Omron Sysmac Studio project 자동화산업기사-고건우_3 (Sysmac Studio 1.53.0.9, StandardProject)

# Controller CPU1: NX102-1020 version 1.33
Units and slaves: 노드1 : NX-ECC203 (E001); 유니트 1 : NX-ID6142-6 (N1); 유니트 2 : NX-OD6121-6 (N2); 유니트 1 : NX-PF0730 (N3); 유니트 2 : NX-ILM400 (N4); 유니트 4 : NX-SID800 (N6); 유니트 5 : NX-SOD400 (N7)
Task PrimaryTask (priority 4, period or condition 2000): Program0

TYPE D_out : UNION
    dw : DWORD;
    b : ARRAY[0..32] OF bool;
END_UNION END_TYPE
TYPE D_in : UNION
    dw : DWORD;
    b : ARRAY[0..32] OF bool;
END_UNION END_TYPE
TYPE U_IO16 : UNION
    W : WORD;
    B : ARRAY[1..32] OF BOOL;
END_UNION END_TYPE
TYPE S_RobotIO : STRUCT
    IO : U_IO16;
END_STRUCT END_TYPE

VAR_GLOBAL
    Bot_Task_Pause : BOOL;  (* 로봇 - 테스크 일시정지; at ECAT://node#[1,2]/Output Bit 32 bits/Output Bit 04 *)
    Discharge_F_SOL : BOOL;  (* at ECAT://node#[1,2]/Output Bit 32 bits/Output Bit 05 *)
    Discharge_R_SS : BOOL;  (* at ECAT://node#[1,1]/Input Bit 32 bits/Input Bit 25 *)
    N1_Input_Bit_26 : BOOL;
    N1_Input_Bit_27 : BOOL;
    N1_Input_Bit_28 : BOOL;
    N1_Input_Bit_29 : BOOL;
    N1_Input_Bit_30 : BOOL;
    N1_Input_Bit_31 : BOOL;
    MotM : WORD;  (* at ECAT://node#2/Command *)
    Vision_Trigger : BOOL;  (* at ECAT://node#4/Line0 Trigger *)
    MotM_Status : WORD;  (* at ECAT://node#2/Status *)
    Robot_Recv : S_RobotIO;
    Robot_Send : S_RobotIO;
    Robot_In : ARRAY[0..237] OF WORD;  (* network input *)
    Robot_Out : ARRAY[0..105] OF WORD;  (* network output *)
END_VAR
VAR_GLOBAL RETAIN
    Bot_IO : ARRAY[1..7] OF WORD := [16#01, 16#02, 16#04, 16#08, 16#10, 16#20, 16#40];
END_VAR
VAR_GLOBAL
    Discharge_R_SOL : BOOL;  (* at ECAT://node#[1,2]/Output Bit 32 bits/Output Bit 06 *)
    Bot_Task_Stop : BOOL;  (* 로봇 - 프로그램 정지; at ECAT://node#[1,2]/Output Bit 32 bits/Output Bit 24 *)
    TWL_R : BOOL;  (* 타워램프 - RED; at ECAT://node#[1,2]/Output Bit 32 bits/Output Bit 20 *)
    TWL_Y : BOOL;  (* 타워램프 - YELLOW; at ECAT://node#[1,2]/Output Bit 32 bits/Output Bit 21 *)
    TWL_G : BOOL;  (* 타워램프 - GREEN; at ECAT://node#[1,2]/Output Bit 32 bits/Output Bit 22 *)
    Bot_Task_ON : BOOL;  (* 로봇 - 태스크 실행; at ECAT://node#[1,2]/Output Bit 32 bits/Output Bit 23 *)
    Vision_SS : BOOL;  (* at ECAT://node#[1,1]/Input Bit 32 bits/Input Bit 19 *)
    Stopper_SS : BOOL;  (* at ECAT://node#[1,1]/Input Bit 32 bits/Input Bit 24 *)
    Magazine_SS : BOOL;  (* at ECAT://node#[1,1]/Input Bit 32 bits/Input Bit 23 *)
    Discharge_F_SS : BOOL;  (* at ECAT://node#[1,1]/Input Bit 32 bits/Input Bit 26 *)
    Bot_Task_Resume : BOOL;  (* 로봇 - 테스크 재개; at ECAT://node#[1,2]/Output Bit 32 bits/Output Bit 13 *)
    Vis_Data : DINT;  (* at ECAT://node#4/Line0 DINT Result Data 0 *)
    H_Count_Val : INT;
    H_Total_Val : INT;
    Robot_DI : S_RobotIO;
    MultiMode_PB : BOOL;
    SingleMode_PB : BOOL;
    Target_Slot_Status : ARRAY[1..6] OF BOOL;
    Stop_PB : BOOL;
    Auto_PB : BOOL;
    Manual_PB : BOOL;
    MotMV_PB : BOOL;
    MotST_PB : BOOL;
    F_SOL_PB : BOOL;
    R_SOL_PB : BOOL;
    Clamp_PB : BOOL;
    UnClamp_PB : BOOL;
    H_Err_Val : INT;
    Auto_Busy : BOOL;
    Manual_Busy : BOOL;
    Pause_PB : BOOL;
    Resume_PB : BOOL;
    Estop_PB : BOOL;
    RST_PB : BOOL;
    gDMemory : WORD;
END_VAR

(* Program Program0: safety or other program stored in binary form, left out *)

PROGRAM Program0
VAR
    i : INT;
    Start : BOOL;
    Vis_ON : BOOL;
    data : INT;
    Sensor_OK : BOOL;
    Pause : BOOL;
    T0 : TON;
    T0TImer : DINT;
    TP0 : TP;
    AT0 : AccumulationTimer;
    Auto : Equipment;
END_VAR
VAR_EXTERNAL
    MotM : WORD;
    Vision_Trigger : BOOL;
    MotM_Status : WORD;
    Magazine_SS : BOOL;
    Discharge_R_SS : BOOL;
    Stopper_SS : BOOL;
    Discharge_F_SS : BOOL;
    Vision_SS : BOOL;
    Vis_Data : DINT;
    Robot_Recv : S_RobotIO;
    Discharge_F_SOL : BOOL;
    Discharge_R_SOL : BOOL;
    Robot_Send : S_RobotIO;
    Bot_Task_Stop : BOOL;
    Bot_Task_ON : BOOL;
    Robot_In : ARRAY[0..237] OF WORD;
    Robot_Out : ARRAY[0..105] OF WORD;
    Bot_Task_Pause : BOOL;
    Bot_Task_Resume : BOOL;
    Bot_IO : ARRAY[1..7] OF WORD;
    H_Count_Val : INT;
    H_Total_Val : INT;
    Robot_DI : S_RobotIO;
    MultiMode_PB : BOOL;
    SingleMode_PB : BOOL;
    Target_Slot_Status : ARRAY[1..6] OF BOOL;
    Stop_PB : BOOL;
    Auto_PB : BOOL;
    Manual_PB : BOOL;
    MotMV_PB : BOOL;
    MotST_PB : BOOL;
    F_SOL_PB : BOOL;
    R_SOL_PB : BOOL;
    Clamp_PB : BOOL;
    UnClamp_PB : BOOL;
    H_Err_Val : INT;
    Auto_Busy : BOOL;
    Manual_Busy : BOOL;
    Pause_PB : BOOL;
    Resume_PB : BOOL;
    Estop_PB : BOOL;
    RST_PB : BOOL;
    TWL_G : BOOL;
    TWL_R : BOOL;
    TWL_Y : BOOL;
END_VAR

(* Section Section0: ladder, written here as Structured Text *)

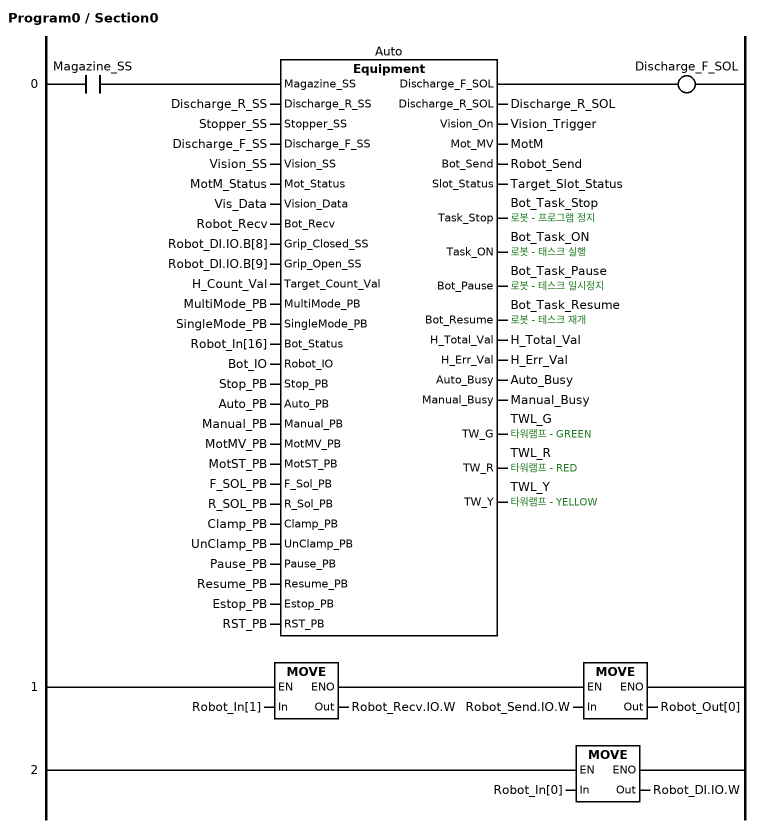
(* Rung 0 *)
Auto(Magazine_SS := Magazine_SS, Discharge_R_SS := Discharge_R_SS, Stopper_SS := Stopper_SS, Discharge_F_SS := Discharge_F_SS, Vision_SS := Vision_SS, Mot_Status := MotM_Status, Vision_Data := Vis_Data, Bot_Recv := Robot_Recv, Grip_Closed_SS := Robot_DI.IO.B[8], Grip_Open_SS := Robot_DI.IO.B[9], Target_Count_Val := H_Count_Val, MultiMode_PB := MultiMode_PB, SingleMode_PB := SingleMode_PB, Bot_Status := Robot_In[16], Robot_IO := Bot_IO, Stop_PB := Stop_PB, Auto_PB := Auto_PB, Manual_PB := Manual_PB, MotMV_PB := MotMV_PB, MotST_PB := MotST_PB, F_Sol_PB := F_SOL_PB, R_Sol_PB := R_SOL_PB, Clamp_PB := Clamp_PB, UnClamp_PB := UnClamp_PB, Pause_PB := Pause_PB, Resume_PB := Resume_PB, Estop_PB := Estop_PB, RST_PB := RST_PB, Discharge_R_SOL => Discharge_R_SOL, Vision_On => Vision_Trigger, Mot_MV => MotM, Bot_Send => Robot_Send, Slot_Status => Target_Slot_Status, Task_Stop => Bot_Task_Stop, Task_ON => Bot_Task_ON, Bot_Pause => Bot_Task_Pause, Bot_Resume => Bot_Task_Resume, H_Total_Val => H_Total_Val, H_Err_Val => H_Err_Val, Auto_Busy => Auto_Busy, Manual_Busy => Manual_Busy, TW_G => TWL_G, TW_R => TWL_R, TW_Y => TWL_Y);
Discharge_F_SOL := Auto.Discharge_F_SOL;
(* Rung 1 *)
Robot_Recv.IO.W := Robot_In[1];
Robot_Out[0] := Robot_Send.IO.W;
(* Rung 2 *)
Robot_DI.IO.W := Robot_In[0];
END_PROGRAM

FUNCTION_BLOCK MPS
VAR
    data : INT;
    T0 : TON;
END_VAR
VAR_INPUT
    MPS_Start : BOOL;
    Discharge_R_SS : BOOL;
    Stopper_SS : BOOL;
END_VAR
VAR_OUTPUT
    Discharge_F_SOL : BOOL;
END_VAR
VAR_INPUT
    Discharge_F_SS : BOOL;
END_VAR
VAR_OUTPUT
    Discharge_R_SOL : BOOL;
END_VAR
VAR_INPUT
    Vision_SS : BOOL;
END_VAR
VAR_OUTPUT
    Vision_On : BOOL;
END_VAR
VAR_INPUT
    Mot_Status : WORD;
END_VAR
VAR_OUTPUT
    MPS_Done : BOOL;
END_VAR
VAR_INPUT
    Cmd_Ack : BOOL;
END_VAR
VAR_OUTPUT
    MPS_Busy : BOOL;
END_VAR
VAR_INPUT
    Vision_Data : DINT;
END_VAR
VAR_OUTPUT
    VIs_NO : DINT;
END_VAR
VAR_IN_OUT
    Mot_MV : WORD;
END_VAR
VAR_INPUT
    Estop_Active : BOOL;
    RST_Active : BOOL;
    Slot_Status : ARRAY[1..6] OF BOOL;
    Pause_Active : BOOL;
END_VAR
VAR
    _e1 : R_TRIG;
    _p2 : BOOL;
    _p3 : BOOL;
END_VAR
(* ladder, written here as Structured Text *)

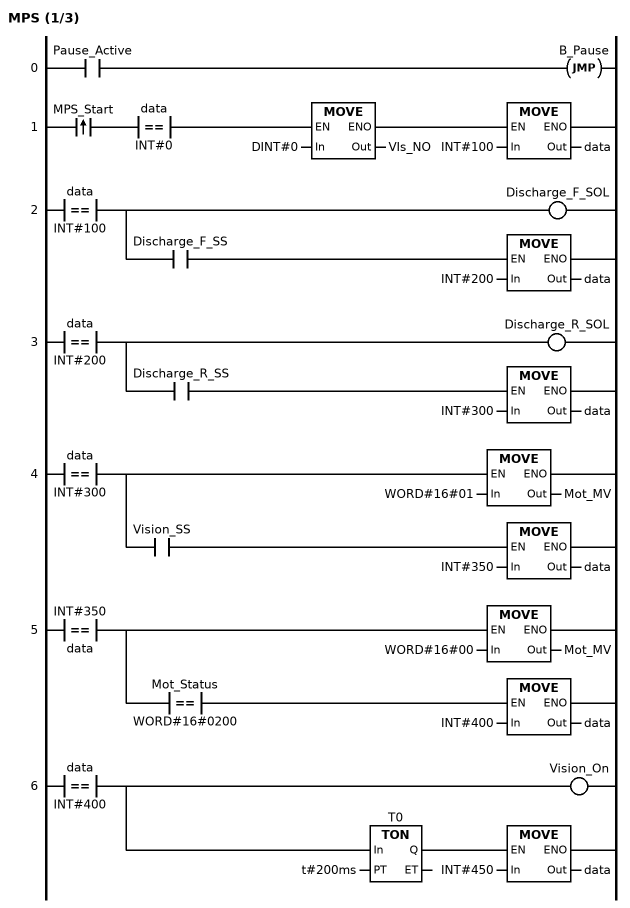
(* Rung 0 *)
IF Pause_Active THEN JMP B_Pause; END_IF;
(* Rung 1 *)
_e1(CLK := MPS_Start);
IF _e1.Q AND (data = INT#0) THEN
    VIs_NO := DINT#0;
    data := INT#100;
END_IF;
(* Rung 2 *)
Discharge_F_SOL := data = INT#100;
IF (data = INT#100) AND Discharge_F_SS THEN data := INT#200; END_IF;
(* Rung 3 *)
Discharge_R_SOL := data = INT#200;
IF (data = INT#200) AND Discharge_R_SS THEN data := INT#300; END_IF;
(* Rung 4 *)
IF data = INT#300 THEN Mot_MV := WORD#16#01; END_IF;
IF (data = INT#300) AND Vision_SS THEN data := INT#350; END_IF;
(* Rung 5 *)
IF INT#350 = data THEN Mot_MV := WORD#16#00; END_IF;
IF (INT#350 = data) AND (Mot_Status = WORD#16#0200) THEN data := INT#400; END_IF;
(* Rung 6 *)
Vision_On := data = INT#400;
T0(In := data = INT#400, PT := t#200ms);
IF T0.Q THEN data := INT#450; END_IF;

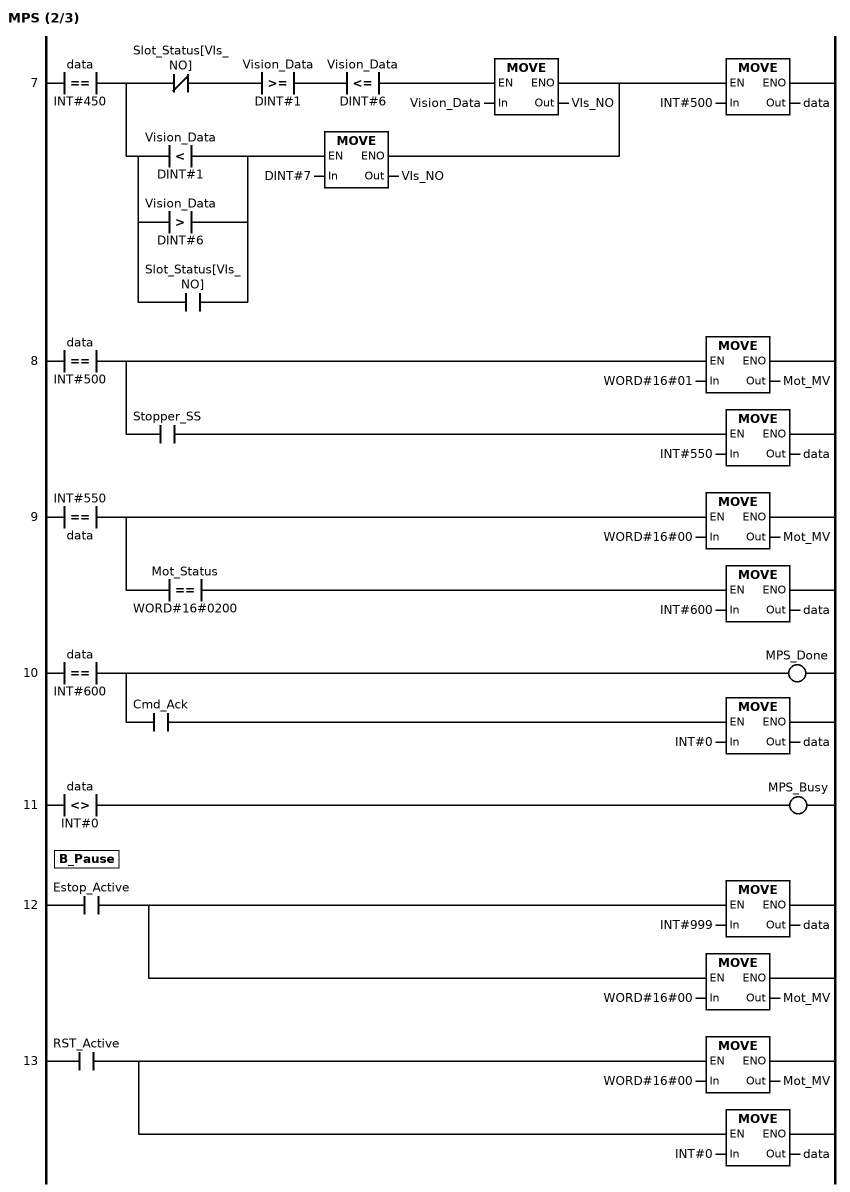
(* Rung 7 *)
_p2 := (data = INT#450) AND NOT Slot_Status[VIs_NO] AND (Vision_Data >= DINT#1) AND (Vision_Data <= DINT#6);
IF _p2 THEN VIs_NO := Vision_Data; END_IF;
_p3 := (data = INT#450) AND ((Vision_Data < DINT#1) OR (Vision_Data > DINT#6) OR Slot_Status[VIs_NO]);
IF _p3 THEN VIs_NO := DINT#7; END_IF;
IF _p2 OR _p3 THEN data := INT#500; END_IF;
(* Rung 8 *)
IF data = INT#500 THEN Mot_MV := WORD#16#01; END_IF;
IF (data = INT#500) AND Stopper_SS THEN data := INT#550; END_IF;
(* Rung 9 *)
IF INT#550 = data THEN Mot_MV := WORD#16#00; END_IF;
IF (INT#550 = data) AND (Mot_Status = WORD#16#0200) THEN data := INT#600; END_IF;
(* Rung 10 *)
MPS_Done := data = INT#600;
IF (data = INT#600) AND Cmd_Ack THEN data := INT#0; END_IF;
(* Rung 11 *)
MPS_Busy := data <> INT#0;
(* Rung 12 *)
B_Pause:
IF Estop_Active THEN
    data := INT#999;
    Mot_MV := WORD#16#00;
END_IF;
(* Rung 13 *)
IF RST_Active THEN
    Mot_MV := WORD#16#00;
    data := INT#0;
END_IF;

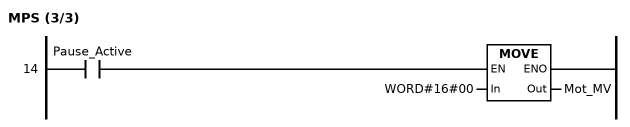
(* Rung 14 *)
IF Pause_Active THEN Mot_MV := WORD#16#00; END_IF;
END_FUNCTION_BLOCK

FUNCTION_BLOCK Robot
VAR
    data : INT;
    T0 : TON;
END_VAR
VAR_INPUT
    Bot_Start : BOOL;
END_VAR
VAR_OUTPUT
    Bot_Done : BOOL;
    Bot_Busy : BOOL;
END_VAR
VAR_IN_OUT
    Slot_Status : ARRAY[1..6] OF BOOL;
END_VAR
VAR_INPUT
    Estop_Active : BOOL;
    RST_Active : BOOL;
    Pause_Active : BOOL;
    Target_Slot_No : DINT;
    MultiMode : BOOL;
END_VAR
VAR_IN_OUT
    Bot_Send : S_RobotIO;
END_VAR
VAR_INPUT
    Bot_Recv : S_RobotIO;
    Bot_Status : WORD;
    Bot_IO : ARRAY[1..7] OF WORD;
END_VAR
VAR_IN_OUT
    H_Total_Val : INT;
    H_Err_Val : INT;
END_VAR
VAR
    _p1 : BOOL;
    _e2 : R_TRIG;
    _e3 : R_TRIG;
END_VAR
(* ladder, written here as Structured Text *)

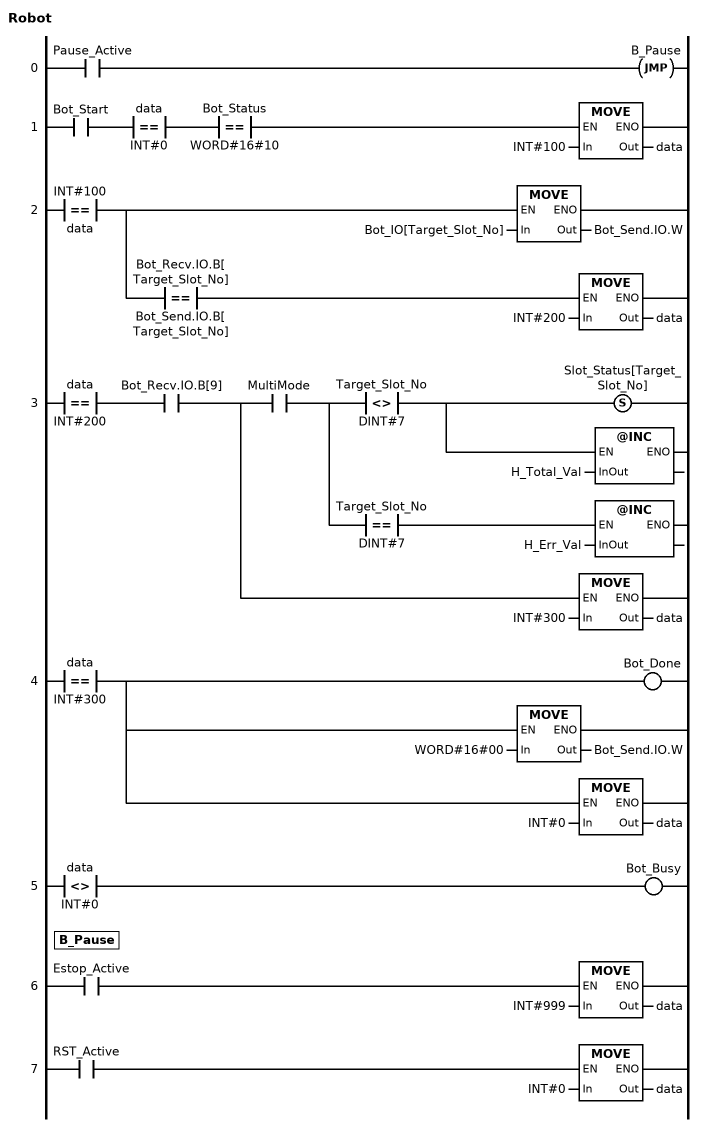
(* Rung 0 *)
IF Pause_Active THEN JMP B_Pause; END_IF;
(* Rung 1 *)
IF Bot_Start AND (data = INT#0) AND (Bot_Status = WORD#16#10) THEN data := INT#100; END_IF;
(* Rung 2 *)
IF INT#100 = data THEN Bot_Send.IO.W := Bot_IO[Target_Slot_No]; END_IF;
IF (INT#100 = data) AND (Bot_Recv.IO.B[Target_Slot_No] = Bot_Send.IO.B[Target_Slot_No]) THEN
    data := INT#200;
END_IF;
(* Rung 3 *)
_p1 := (data = INT#200) AND Bot_Recv.IO.B[9] AND MultiMode;
IF _p1 AND (Target_Slot_No <> DINT#7) THEN Slot_Status[Target_Slot_No] := TRUE; END_IF;
_e2(CLK := _p1 AND (Target_Slot_No <> DINT#7));
IF _e2.Q THEN INC(InOut := H_Total_Val); END_IF;
_e3(CLK := _p1 AND (Target_Slot_No = DINT#7));
IF _e3.Q THEN INC(InOut := H_Err_Val); END_IF;
IF (data = INT#200) AND Bot_Recv.IO.B[9] THEN data := INT#300; END_IF;
(* Rung 4 *)
Bot_Done := data = INT#300;
IF data = INT#300 THEN
    Bot_Send.IO.W := WORD#16#00;
    data := INT#0;
END_IF;
(* Rung 5 *)
Bot_Busy := data <> INT#0;
(* Rung 6 *)
B_Pause:
IF Estop_Active THEN data := INT#999; END_IF;
(* Rung 7 *)
IF RST_Active THEN data := INT#0; END_IF;
END_FUNCTION_BLOCK

FUNCTION_BLOCK Equipment
VAR
    Conveyor : MPS;
    Doosan : Robot;
    Bot_Busy : BOOL;
    Mps_Done : BOOL;
    Mps_Busy : BOOL;
    Vis_No : DINT;
    Bot_Done : BOOL;
    Single_Busy : BOOL;
    Multi_Busy : BOOL;
    C0 : CTU;
    Estop_Active : BOOL;
    RST_Active : BOOL;
    Pause_Active : BOOL;
    Retry : BOOL;
    CTU_RST : BOOL;
    T0 : TON;
    T1 : TON;
    T2 : TON;
    RST_On : BOOL;
    RST_Discharge_R_SOL : BOOL;
    MPS_Discharge_R_SOL : BOOL;
    Stop_Active : BOOL;
    Manual : Passive;
    Manu_Discharge_F_SOL : BOOL;
    Manu_Discharge_R_SOL : BOOL;
    Manu_TWL_G : BOOL;
    MPS_Discharge_F_SOL : BOOL;
    T3 : TON;
    Ready : BOOL;
    Pulse_Pause : BOOL;
    Pause_Eq : BOOL;
END_VAR
VAR_INPUT
    Magazine_SS : BOOL;
    Discharge_R_SS : BOOL;
    Stopper_SS : BOOL;
    Discharge_F_SS : BOOL;
    Vision_SS : BOOL;
    Mot_Status : WORD;
    Vision_Data : DINT;
END_VAR
VAR_OUTPUT
    Discharge_F_SOL : BOOL;
    Discharge_R_SOL : BOOL;
    Vision_On : BOOL;
    Mot_MV : WORD;
END_VAR
VAR_INPUT
    Bot_Recv : S_RobotIO;
END_VAR
VAR_OUTPUT
    Bot_Send : S_RobotIO;
END_VAR
VAR_INPUT
    Grip_Closed_SS : BOOL;
    Grip_Open_SS : BOOL;
END_VAR
VAR_OUTPUT
    Slot_Status : ARRAY[1..6] OF BOOL;
    Task_Stop : BOOL;
END_VAR
VAR_INPUT
    Target_Count_Val : INT;
    MultiMode_PB : BOOL;
    SingleMode_PB : BOOL;
END_VAR
VAR_OUTPUT
    Task_ON : BOOL;
END_VAR
VAR_INPUT
    Bot_Status : WORD;
END_VAR
VAR_OUTPUT
    Bot_Pause : BOOL;
    Bot_Resume : BOOL;
END_VAR
VAR_INPUT
    Robot_IO : ARRAY[1..7] OF WORD;
END_VAR
VAR_OUTPUT
    H_Total_Val : INT;
END_VAR
VAR_INPUT
    Stop_PB : BOOL;
    Auto_PB : BOOL;
    Manual_PB : BOOL;
    MotMV_PB : BOOL;
    MotST_PB : BOOL;
    F_Sol_PB : BOOL;
    R_Sol_PB : BOOL;
    Clamp_PB : BOOL;
    UnClamp_PB : BOOL;
END_VAR
VAR_OUTPUT
    H_Err_Val : INT;
    Auto_Busy : BOOL;
    Manual_Busy : BOOL;
END_VAR
VAR_INPUT
    Pause_PB : BOOL;
    Resume_PB : BOOL;
    Estop_PB : BOOL;
    RST_PB : BOOL;
END_VAR
VAR_OUTPUT
    TW_G : BOOL;
    TW_R : BOOL;
    TW_Y : BOOL;
END_VAR
VAR
    _e1 : R_TRIG;
    _p2 : BOOL;
    _e3 : F_TRIG;
    _e4 : R_TRIG;
    _e5 : R_TRIG;
END_VAR
(* ladder, written here as Structured Text *)

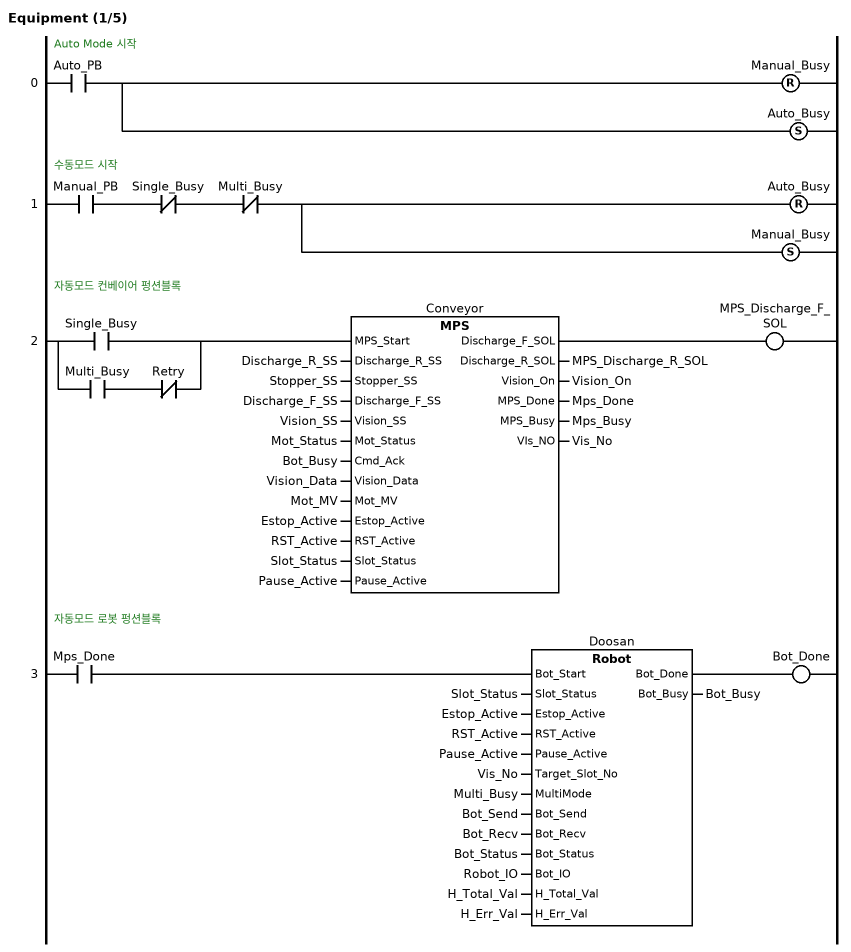
(* Rung 0: Auto Mode 시작 *)
IF Auto_PB THEN
    Manual_Busy := FALSE;
    Auto_Busy := TRUE;
END_IF;
(* Rung 1: 수동모드 시작 *)
IF Manual_PB AND NOT Single_Busy AND NOT Multi_Busy THEN
    Auto_Busy := FALSE;
    Manual_Busy := TRUE;
END_IF;
(* Rung 2: 자동모드 컨베이어 펑션블록 *)
Conveyor(MPS_Start := Single_Busy OR (Multi_Busy AND NOT Retry), Discharge_R_SS := Discharge_R_SS, Stopper_SS := Stopper_SS, Discharge_F_SS := Discharge_F_SS, Vision_SS := Vision_SS, Mot_Status := Mot_Status, Cmd_Ack := Bot_Busy, Vision_Data := Vision_Data, Mot_MV := Mot_MV, Estop_Active := Estop_Active, RST_Active := RST_Active, Slot_Status := Slot_Status, Pause_Active := Pause_Active, Discharge_R_SOL => MPS_Discharge_R_SOL, Vision_On => Vision_On, MPS_Done => Mps_Done, MPS_Busy => Mps_Busy, VIs_NO => Vis_No);
MPS_Discharge_F_SOL := Conveyor.Discharge_F_SOL;
(* Rung 3: 자동모드 로봇 펑션블록 *)
Doosan(Bot_Start := Mps_Done, Slot_Status := Slot_Status, Estop_Active := Estop_Active, RST_Active := RST_Active, Pause_Active := Pause_Active, Target_Slot_No := Vis_No, MultiMode := Multi_Busy, Bot_Send := Bot_Send, Bot_Recv := Bot_Recv, Bot_Status := Bot_Status, Bot_IO := Robot_IO, H_Total_Val := H_Total_Val, H_Err_Val := H_Err_Val, Bot_Busy => Bot_Busy);
Bot_Done := Doosan.Bot_Done;

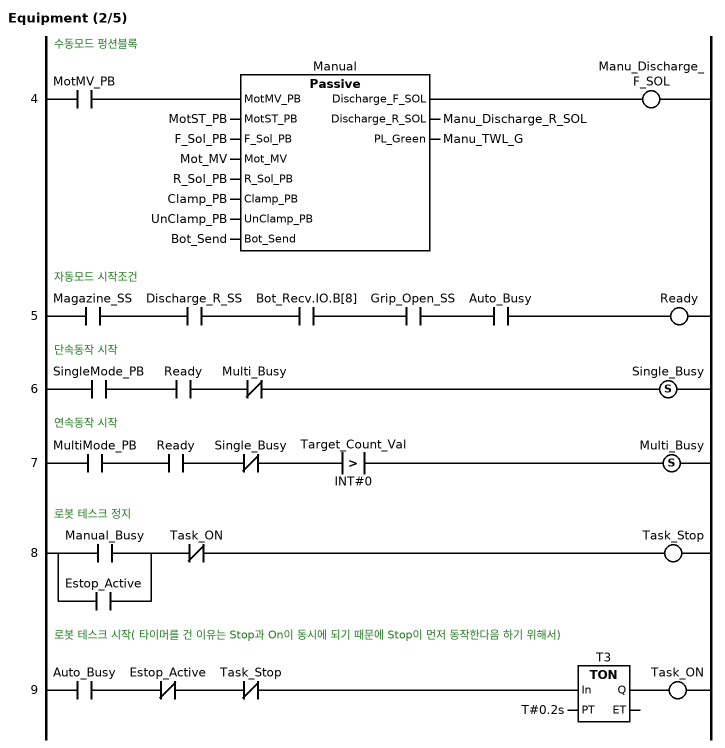
(* Rung 4: 수동모드 펑션블록 *)
Manual(MotMV_PB := MotMV_PB, MotST_PB := MotST_PB, F_Sol_PB := F_Sol_PB, Mot_MV := Mot_MV, R_Sol_PB := R_Sol_PB, Clamp_PB := Clamp_PB, UnClamp_PB := UnClamp_PB, Bot_Send := Bot_Send, Discharge_R_SOL => Manu_Discharge_R_SOL, PL_Green => Manu_TWL_G);
Manu_Discharge_F_SOL := Manual.Discharge_F_SOL;
(* Rung 5: 자동모드 시작조건 *)
Ready := Magazine_SS AND Discharge_R_SS AND Bot_Recv.IO.B[8] AND Grip_Open_SS AND Auto_Busy;
(* Rung 6: 단속동작 시작 *)
IF SingleMode_PB AND Ready AND NOT Multi_Busy THEN Single_Busy := TRUE; END_IF;
(* Rung 7: 연속동작 시작 *)
IF MultiMode_PB AND Ready AND NOT Single_Busy AND (Target_Count_Val > INT#0) THEN
    Multi_Busy := TRUE;
END_IF;
(* Rung 8: 로봇 테스크 정지 *)
Task_Stop := (Manual_Busy OR Estop_Active) AND NOT Task_ON;
(* Rung 9: 로봇 테스크 시작( 타이머를 건 이유는 Stop과 On이 동시에 되기 때문에 Stop이 먼저 동작한다음 하기 위해서) *)
T3(In := Auto_Busy AND NOT Estop_Active AND NOT Task_Stop, PT := T#0.2s);
Task_ON := T3.Q;

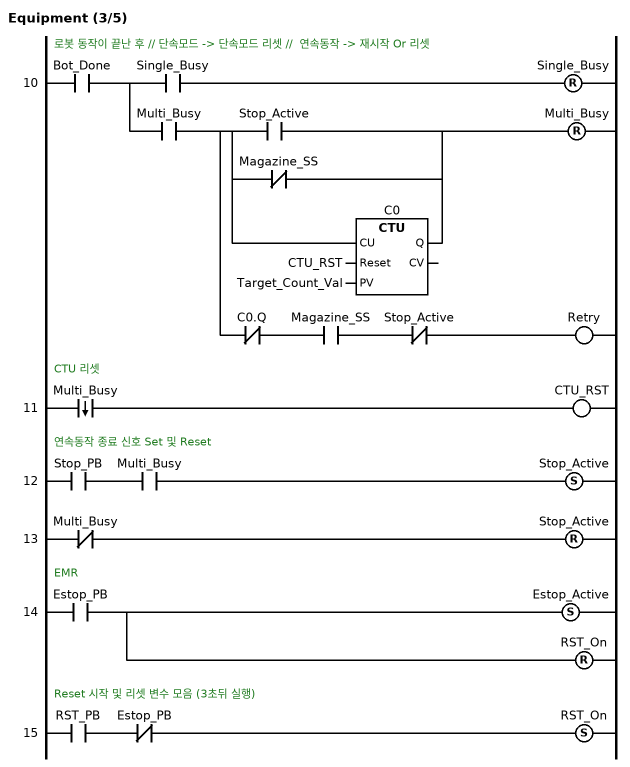
(* Rung 10: 로봇 동작이 끝난 후 // 단속모드 -> 단속모드 리셋 //  연속동작 -> 재시작 Or 리셋 *)
IF Bot_Done AND Single_Busy THEN Single_Busy := FALSE; END_IF;
_e1(CLK := Bot_Done AND Multi_Busy);
C0(CU := _e1.Q, Reset := CTU_RST, PV := Target_Count_Val);
_p2 := Bot_Done AND Multi_Busy;
IF (Bot_Done AND Multi_Busy AND (Stop_Active OR NOT Magazine_SS)) OR C0.Q THEN
    Multi_Busy := FALSE;
END_IF;
Retry := _p2 AND NOT C0.Q AND Magazine_SS AND NOT Stop_Active;
(* Rung 11: CTU 리셋 *)
_e3(CLK := Multi_Busy);
CTU_RST := _e3.Q;
(* Rung 12: 연속동작 종료 신호 Set 및 Reset *)
IF Stop_PB AND Multi_Busy THEN Stop_Active := TRUE; END_IF;
(* Rung 13 *)
IF NOT Multi_Busy THEN Stop_Active := FALSE; END_IF;
(* Rung 14: EMR *)
IF Estop_PB THEN
    Estop_Active := TRUE;
    RST_On := FALSE;
END_IF;
(* Rung 15: Reset 시작 및 리셋 변수 모음 (3초뒤 실행) *)
IF RST_PB AND NOT Estop_PB THEN RST_On := TRUE; END_IF;

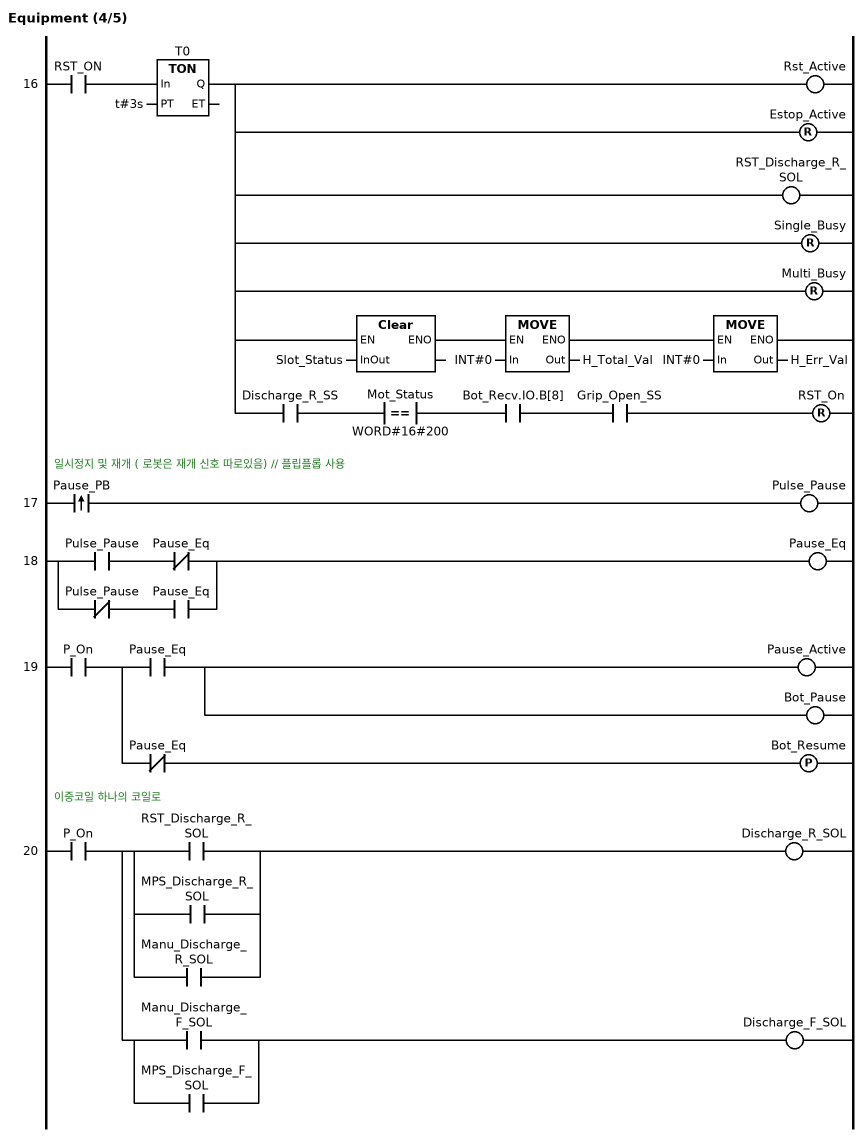
(* Rung 16 *)
T0(In := RST_ON, PT := t#3s);
Rst_Active := T0.Q;
IF T0.Q THEN Estop_Active := FALSE; END_IF;
RST_Discharge_R_SOL := T0.Q;
IF T0.Q THEN
    Single_Busy := FALSE;
    Multi_Busy := FALSE;
    Clear(InOut := Slot_Status);
    H_Total_Val := INT#0;
    H_Err_Val := INT#0;
END_IF;
IF T0.Q AND Discharge_R_SS AND (Mot_Status = WORD#16#200) AND Bot_Recv.IO.B[8] AND Grip_Open_SS THEN
    RST_On := FALSE;
END_IF;
(* Rung 17: 일시정지 및 재개 ( 로봇은 재개 신호 따로있음) // 플립플롭 사용 *)
_e4(CLK := Pause_PB);
Pulse_Pause := _e4.Q;
(* Rung 18 *)
Pause_Eq := (Pulse_Pause AND NOT Pause_Eq) OR (NOT Pulse_Pause AND Pause_Eq);
(* Rung 19 *)
Pause_Active := P_On AND Pause_Eq;
Bot_Pause := P_On AND Pause_Eq;
_e5(CLK := P_On AND NOT Pause_Eq);
Bot_Resume := _e5.Q;
(* Rung 20: 이중코일 하나의 코일로 *)
Discharge_R_SOL := P_On AND (RST_Discharge_R_SOL OR MPS_Discharge_R_SOL OR Manu_Discharge_R_SOL);
Discharge_F_SOL := P_On AND (Manu_Discharge_F_SOL OR MPS_Discharge_F_SOL);

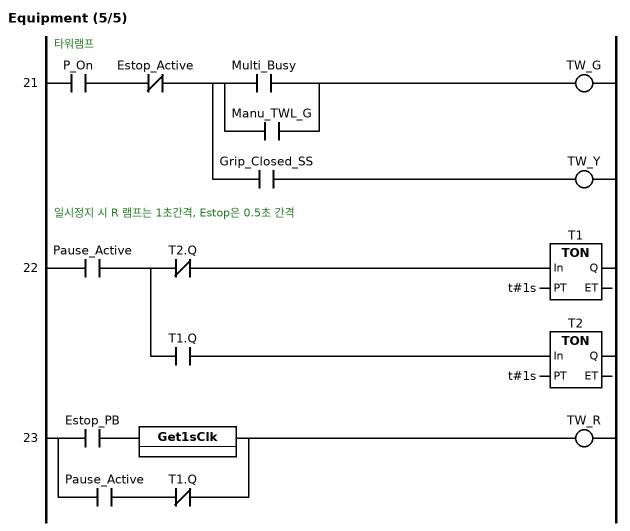
(* Rung 21: 타워램프 *)
TW_G := P_On AND NOT Estop_Active AND (Multi_Busy OR Manu_TWL_G);
TW_Y := P_On AND NOT Estop_Active AND Grip_Closed_SS;
(* Rung 22: 일시정지 시 R 램프는 1초간격, Estop은 0.5초 간격 *)
T1(In := Pause_Active AND NOT T2.Q, PT := t#1s);
T2(In := Pause_Active AND T1.Q, PT := t#1s);
(* Rung 23 *)
TW_R := (Estop_PB AND Get1sClk()) OR (Pause_Active AND NOT T1.Q);
END_FUNCTION_BLOCK

FUNCTION_BLOCK Passive
VAR_INPUT
    MotMV_PB : BOOL;
    MotST_PB : BOOL;
    F_Sol_PB : BOOL;
END_VAR
VAR_OUTPUT
    Discharge_F_SOL : BOOL;
    Discharge_R_SOL : BOOL;
END_VAR
VAR_IN_OUT
    Mot_MV : WORD;
END_VAR
VAR_INPUT
    R_Sol_PB : BOOL;
END_VAR
VAR_OUTPUT
    PL_Green : BOOL;
END_VAR
VAR_INPUT
    Clamp_PB : BOOL;
    UnClamp_PB : BOOL;
END_VAR
VAR_IN_OUT
    Bot_Send : S_RobotIO;
END_VAR
(* ladder, written here as Structured Text *)

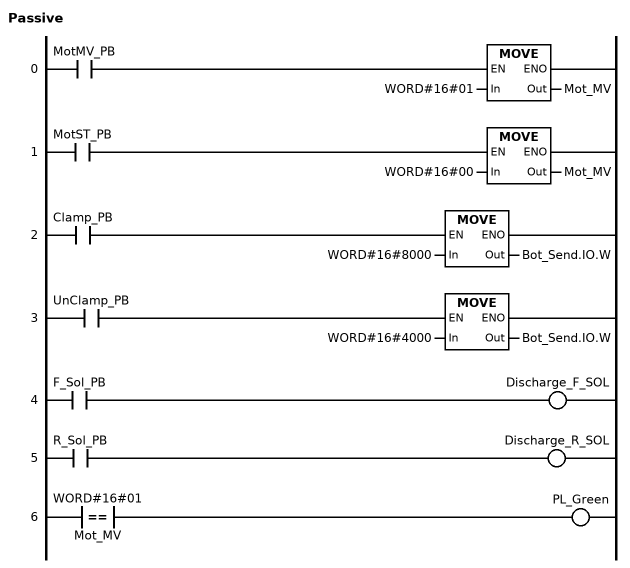
(* Rung 0 *)
IF MotMV_PB THEN Mot_MV := WORD#16#01; END_IF;
(* Rung 1 *)
IF MotST_PB THEN Mot_MV := WORD#16#00; END_IF;
(* Rung 2 *)
IF Clamp_PB THEN Bot_Send.IO.W := WORD#16#8000; END_IF;
(* Rung 3 *)
IF UnClamp_PB THEN Bot_Send.IO.W := WORD#16#4000; END_IF;
(* Rung 4 *)
Discharge_F_SOL := F_Sol_PB;
(* Rung 5 *)
Discharge_R_SOL := R_Sol_PB;
(* Rung 6 *)
PL_Green := WORD#16#01 = Mot_MV;
END_FUNCTION_BLOCK

# Device HMI_NA5_0 (NA): not converted